(* IEC 61131-3 sources: Test-Git_ESME26/TestProgettoESME_26.fbsproj/PacDriveLib Migration/Motion/MultiCam/PDL_FB_MultiCam.fb.st^/SetOutputs, 5 files *)

(* ---- InWindowMode.meth.st ---- *)
METHOD PRIVATE InWindowMode : BOOL
//only in ws mode ___CamShowCamPosition
//sets output q_xInWSWindow
VAR_INPUT
END_VAR
VAR
END_VAR

InWindowMode := TRUE;

lrPositionY2:= i_ifDrive.lrPosition;

IF stActiveMultiCamData.lrYPeriod <> 0 THEN
	lrYPeriode := stActiveMultiCamData.lrYPeriod;
END_IF

CASE iq_stExt.etInWindowMode OF

	PDL_ET_MultiCamWsMode.StoredCamMoveAlwaysNoPositionCheck,
	PDL_ET_MultiCamWsMode.StoredCamMoveToCamPositonInWsWindow,
	PDL_ET_MultiCamWsMode.NewCamMoveAlwaysNoPositionCheck,
	PDL_ET_MultiCamWsMode.NewCamMoveToCamPositonInWsWindow:

		IF NOT iq_stExt.xNoModuloSlaveAtStart THEN
			IF ABS(lrYStart - lrPositionY2) <= i_lrWSWindow THEN
				q_xInWSWindow := TRUE;

			(* pos. Periode *)
			ELSIF lrYPeriode > 0 AND lrYStart >= lrPositionY2 AND ABS(lrPositionY2 + lrYPeriode - lrYStart) <= i_lrWSWindow THEN
				q_xInWSWindow := TRUE;
			ELSIF lrYPeriode > 0 AND lrYStart < lrPositionY2 AND ABS(lrYStart + lrYPeriode - lrPositionY2) <= i_lrWSWindow THEN
				q_xInWSWindow := TRUE;

			(* neg. Periode *)
			ELSIF lrYPeriode < 0 AND lrYStart <= lrPositionY2 AND ABS(lrYStart - lrPositionY2 - lrYPeriode) <= i_lrWSWindow THEN
				q_xInWSWindow:= TRUE;
			ELSIF lrYPeriode < 0 AND lrYStart > lrPositionY2 AND ABS(lrPositionY2 - lrYPeriode - lrYStart) <= i_lrWSWindow THEN
				q_xInWSWindow := TRUE;
			ELSE
				q_xInWSWindow := FALSE;
			END_IF
		ELSE
			IF ABS(lrYStart - lrPositionY2) <= i_lrWSWindow THEN
				q_xInWSWindow := TRUE;
			ELSE
				q_xInWSWindow := FALSE;
			END_IF
		END_IF

	PDL_ET_MultiCamWsMode.StoredCamMoveForwardToCamPositon,
	PDL_ET_MultiCamWsMode.StoredCamMoveBackwardToCamPosition,
	PDL_ET_MultiCamWsMode.NewCamMoveForwardToCamPositon,
	PDL_ET_MultiCamWsMode.NewCamMoveBackwardToCamPosition:

		IF  iq_stExt.xInWindowCheckwithoutLimits THEN
			IF ABS(lrYStart - lrPositionY2) <= i_lrWSWindow THEN
				q_xInWSWindow := TRUE;

			(* pos. Periode *)
			ELSIF lrYPeriode > 0 AND lrYStart >= lrPositionY2 AND ABS(lrPositionY2 + lrYPeriode - lrYStart) <= i_lrWSWindow THEN
				q_xInWSWindow := TRUE;
			ELSIF lrYPeriode > 0 AND lrYStart < lrPositionY2 AND ABS(lrYStart + lrYPeriode - lrPositionY2) <= i_lrWSWindow THEN
				q_xInWSWindow := TRUE;

			(* neg. Periode *)
			ELSIF lrYPeriode < 0 AND lrYStart <= lrPositionY2 AND ABS(lrYStart - lrPositionY2 - lrYPeriode) <= i_lrWSWindow THEN
				q_xInWSWindow := TRUE;
			ELSIF lrYPeriode < 0 AND lrYStart > lrPositionY2 AND ABS(lrPositionY2 - lrYPeriode - lrYStart) <= i_lrWSWindow THEN
				q_xInWSWindow := TRUE;
			ELSE
				q_xInWSWindow := FALSE;
			END_IF
		ELSE
			IF ABS(lrYStart - lrPositionY2) <= i_lrWSWindow THEN
				q_xInWSWindow := TRUE;
			ELSE
				q_xInWSWindow := FALSE;
			END_IF
		END_IF

ELSE
	q_xInWSWindow := FALSE;
END_CASE

(* ---- SetActualCamData.meth.st ---- *)
METHOD PRIVATE SetActualCamData : BOOL
VAR_INPUT
END_VAR

//set values
q_stActualCamData.diProfileId	:= -1;
q_stActualCamData.lrXOffset		:= stActiveMultiCamData.astCamPoint[0].lrX;
q_stActualCamData.lrYOffset		:= stActiveMultiCamData.astCamPoint[0].lrY;
q_stActualCamData.lrXFactor		:=  stActiveMultiCamData.astCamPoint[stActiveMultiCamData.diNumberOfCamPoints-1].lrX
								  - stActiveMultiCamData.astCamPoint[0].lrX;

MOIN.FC_CamBounds(	i_stCamTableID		:= stActiveMultiCamData,
					i_lrMasterVelMax	:= 0,
					i_lrMasterAccMax	:= 0,
					i_lrMasterScaling	:= 1,
					i_lrSlaveScaling	:= 1,
					q_lrMaxPosition		=> q_stActualCamData.lrYFactor
					);

q_stActualCamData.diUserTableId	:= stActiveMultiCamData.diUserTableId;

lrYPeriode := stActiveMultiCamData.lrYPeriod;
lrXPeriode := stActiveMultiCamData.astCamPoint[stActiveMultiCamData.diNumberOfCamPoints-1].lrX - stActiveMultiCamData.astCamPoint[0].lrX;

(* ---- SetDiagOutput.meth.st ---- *)
METHOD PRIVATE SetDiagOutput : BOOL
VAR_INPUT
	i_etDiag	: GD.ET_Diag;
	i_etDiagExt	: PDL_ET_DiagExt;
	i_sMsg		: STRING[80];
END_VAR
VAR
END_VAR

IF i_etDiag <> GD.ET_Diag.Ok THEN
	q_xReady := FALSE;
END_IF

IF q_etDiag = GD.ET_Diag.OK OR i_etDiagExt = PDL_ET_DiagExt.Disabled THEN
	q_etDiag := i_etDiag;
	q_etDiagExt := i_etDiagExt;
	q_sMsg := i_sMsg;

	IF(i_etDiag = GD.ET_Diag.Ok) AND (THIS^.fbLoggerPoint.etLogLevel >= APL.ET_LogLevel.StatusMessage) THEN
		THIS^.fbLoggerPoint.AddLogEntry(	i_etLogLevel	:= APL.ET_LogLevel.StatusMessage,
											i_etDiag		:= q_etDiag,
											i_udiDiagExt	:= q_etDiagExt,
											i_sMessage		:= SE_CTBX.FC_MultiConcat(	i_sString1	:= Standard.CONCAT('ET_Diag: ', GD.FC_EtDiagToString(q_etDiag)),
																						i_sString2	:= Standard.CONCAT(' ET_DiagExt: ', PDL_FC_EtDiagExtToString(q_etDiagExt)),
																						i_sString3	:= Standard.CONCAT(' sMsg: ', q_sMsg),
																						i_sString4	:= '')
										);

	ELSIF(i_etDiag = GD.ET_Diag.UnexpectedProgramBehavior) AND (THIS^.fbLoggerPoint.etLogLevel >= APL.ET_LogLevel.CriticalException) THEN
		THIS^.fbLoggerPoint.AddLogEntry(	i_etLogLevel	:= APL.ET_LogLevel.CriticalException,
											i_etDiag		:= q_etDiag,
											i_udiDiagExt	:= q_etDiagExt,
											i_sMessage		:= SE_CTBX.FC_MultiConcat(	i_sString1	:= Standard.CONCAT('ET_Diag: ', GD.FC_EtDiagToString(q_etDiag)),
																						i_sString2	:= Standard.CONCAT(' ET_DiagExt: ', PDL_FC_EtDiagExtToString(q_etDiagExt)),
																						i_sString3	:= Standard.CONCAT(' sMsg: ', q_sMsg),
																						i_sString4	:= '')
										);

	ELSIF(i_etDiag <> GD.ET_Diag.Ok) AND (THIS^.fbLoggerPoint.etLogLevel >= APL.ET_LogLevel.Exception) THEN
		THIS^.fbLoggerPoint.AddLogEntry(	i_etLogLevel	:= APL.ET_LogLevel.Exception,
											i_etDiag		:= q_etDiag,
											i_udiDiagExt	:= q_etDiagExt,
											i_sMessage		:= SE_CTBX.FC_MultiConcat(	i_sString1	:= Standard.CONCAT('ET_Diag: ', GD.FC_EtDiagToString(q_etDiag)),
																						i_sString2	:= Standard.CONCAT(' ET_DiagExt: ', PDL_FC_EtDiagExtToString(q_etDiagExt)),
																						i_sString3	:= Standard.CONCAT(' sMsg: ', q_sMsg),
																						i_sString4	:= '')
										);
	END_IF
END_IF

(* ---- SetInWsWindow.meth.st ---- *)
METHOD PRIVATE SetInWsWindow : BOOL
VAR_INPUT
	i_xCheckModulo			: BOOL;
END_VAR

IF 	i_xCheckModulo
THEN
	IF ABS(lrYStart - q_lrPositionY) <= i_lrWSWindow THEN
		q_xInWSWindow := TRUE;
	(* pos. Periode *)
	ELSIF lrYPeriode > 0 AND lrYStart >= q_lrPositionY AND q_lrPositionY + lrYPeriode - lrYStart <= i_lrWSWindow THEN
		q_xInWSWindow := TRUE;
	ELSIF lrYPeriode > 0 AND lrYStart < q_lrPositionY AND lrYStart + lrYPeriode - q_lrPositionY <= i_lrWSWindow THEN
		q_xInWSWindow := TRUE;
	(* neg. Periode *)
	ELSIF lrYPeriode < 0 AND lrYStart <= q_lrPositionY AND lrYStart - q_lrPositionY - lrYPeriode <= i_lrWSWindow THEN
		q_xInWSWindow := TRUE;
	ELSIF lrYPeriode < 0 AND lrYStart > q_lrPositionY AND q_lrPositionY - lrYPeriode - lrYStart <= i_lrWSWindow THEN
		q_xInWSWindow := TRUE;
	ELSE
		q_xInWSWindow := FALSE;
	END_IF
ELSE
	IF ABS(lrYStart - q_lrPositionY) <= i_lrWSWindow THEN
		q_xInWSWindow := TRUE;
	ELSE
		q_xInWSWindow := FALSE;
	END_IF
END_IF

(* ---- SetXHighEnd_XLowEnd.meth.st ---- *)
METHOD PRIVATE SetXHighEnd_XLowEnd : BOOL
VAR_INPUT
END_VAR
VAR
END_VAR

SetXHighEnd_XLowEnd := TRUE;

IF iq_stExt.lrXEndWidth > 0 THEN
	q_xXHighEnd:= (q_lrPositionX >= stActiveMultiCamData.astCamPoint[stActiveMultiCamData.diNumberOfCamPoints-1].lrX   -  iq_stExt.lrXEndWidth);
	q_xXLowEnd:= (q_lrPositionX <= stActiveMultiCamData.astCamPoint[0].lrX +  iq_stExt.lrXEndWidth);

ELSE
(* Set q_xXHighEnd *)
	IF NOT q_xXHighEnd AND lrVelocityX > LREAL#0.0 THEN
		lrXHighEndWidth := lrTSwitch * ABS(lrVelocityX);
		q_xXHighEnd	:= (q_lrPositionX >= stActiveMultiCamData.astCamPoint[stActiveMultiCamData.diNumberOfCamPoints-1].lrX   - lrXHighEndWidth);
	END_IF

(* Set q_xXLowEnd *)
	IF NOT q_xXLowEnd AND lrVelocityX < LREAL#0.0 THEN
		lrXLowEndWidth := lrTSwitch * ABS(lrVelocityX);
		q_xXLowEnd	:= (q_lrPositionX <= stActiveMultiCamData.astCamPoint[0].lrX + lrXLowEndWidth);
	END_IF

(* Reset q_xXHighEnd pos. direction *)
	IF    q_lrPositionX < (stActiveMultiCamData.astCamPoint[stActiveMultiCamData.diNumberOfCamPoints-1].lrX   - lrXHighEndWidth)
	  AND lrVelocityX > LREAL#0.0
	THEN
		q_xXHighEnd := FALSE;
	END_IF

(* Reset q_xXHighEnd neg. direction *)
	IF q_xXLowEnd AND lrVelocityX < LREAL#0.0
	THEN
		q_xXHighEnd := FALSE;
	END_IF

(* Reset q_xXLowEnd neg. direction *)
	IF    q_lrPositionX > (stActiveMultiCamData.astCamPoint[0].lrX + lrXLowEndWidth)
	  AND lrVelocityX < LREAL#0.0
	THEN
		q_xXLowEnd := FALSE;
	END_IF

(* Reset q_xXLowEnd pos. direction *)
	IF    q_xXHighEnd
	  AND lrVelocityX > LREAL#0.0
	THEN
		q_xXLowEnd := FALSE;
	END_IF
END_IF
